// SIMATIC S7-200 project (STEP 7-Micro/WIN), CPU 224 CN REL 02.01

SYMBOL_TABLE USUARIO1
SF1              I0.0     // Sensor optico
SM3              I0.1     // Sensor magnetico de la Pinza
SM2              I0.2     // Sensor magnetico extendido cilindro horizontal
SM1              I0.3     // Sensor magnetico retraido cilindro horizontal
SM4              I0.4     // Sensor magnetico retraido cilindro de compresion
SM5              I0.5     // Sensor magnetico extendido cilindro de compresion
SB_2             I1.2     // Pulsador de paro
SB_1             I1.3     // Pulsador de marcha
QS               I1.4     // Zeta de emergencia
SA               I1.5     // Selector de modo
KV2              Q0.0     // Cilindro de la pinza
KV1              Q0.2     // Cilindro neumatico horizontal
KV3              Q0.3     // Cilindro neumatico de compresion
HL1              Q0.7     // Piloto indicador de parada
HL2              Q1.0     // Piloto indicador de marcha
HL3              Q1.1     // Piloto indicador de emergencia
E0               M0.0     // Estado 0
E1               M0.1     // Estado 1
E2               M0.2     // Estado 2
E3               M0.3     // Estado 3
E4               M0.4     // Estado 4
E5               M0.5     // Estado 5
E6               M0.6     // Estado 6
E7               M0.7     // Estado 7
EP               M1.0     // Estado de parada
EM               M1.1     // Estado de emergencia
END_SYMBOL_TABLE

ORGANIZATION_BLOCK PRINCIPAL:OB1
TITLE=COMENTARIOS DEL PROGRAMA
BEGIN
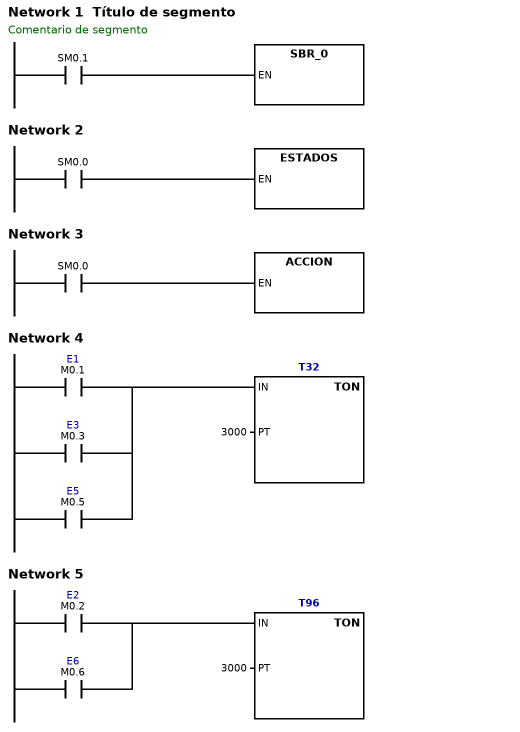
Network 1 // Título de segmento
// Comentario de segmento
LD     SM0.1
CALL   SBR_0:SBR0
Network 2
LD     SM0.0
CALL   ESTADOS:SBR1
Network 3
LD     SM0.0
CALL   ACCION:SBR2
Network 4
LD     E1:M0.1
O      E3:M0.3
O      E5:M0.5
TON    T32, 3000
Network 5
LD     E2:M0.2
O      E6:M0.6
TON    T96, 3000
END_ORGANIZATION_BLOCK

SUBROUTINE_BLOCK SBR_0:SBR0
TITLE=COMENTARIOS DE LA SUBRUTINA
BEGIN
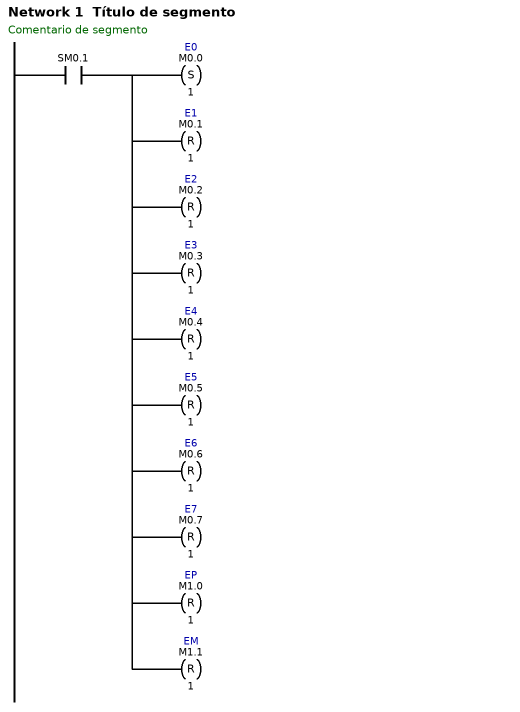
Network 1 // Título de segmento
// Comentario de segmento
LD     SM0.1
S      E0:M0.0, 1
R      E1:M0.1, 1
R      E2:M0.2, 1
R      E3:M0.3, 1
R      E4:M0.4, 1
R      E5:M0.5, 1
R      E6:M0.6, 1
R      E7:M0.7, 1
R      EP:M1.0, 1
R      EM:M1.1, 1
END_SUBROUTINE_BLOCK

SUBROUTINE_BLOCK ESTADOS:SBR1
TITLE=COMENTARIOS DE LA SUBRUTINA
BEGIN
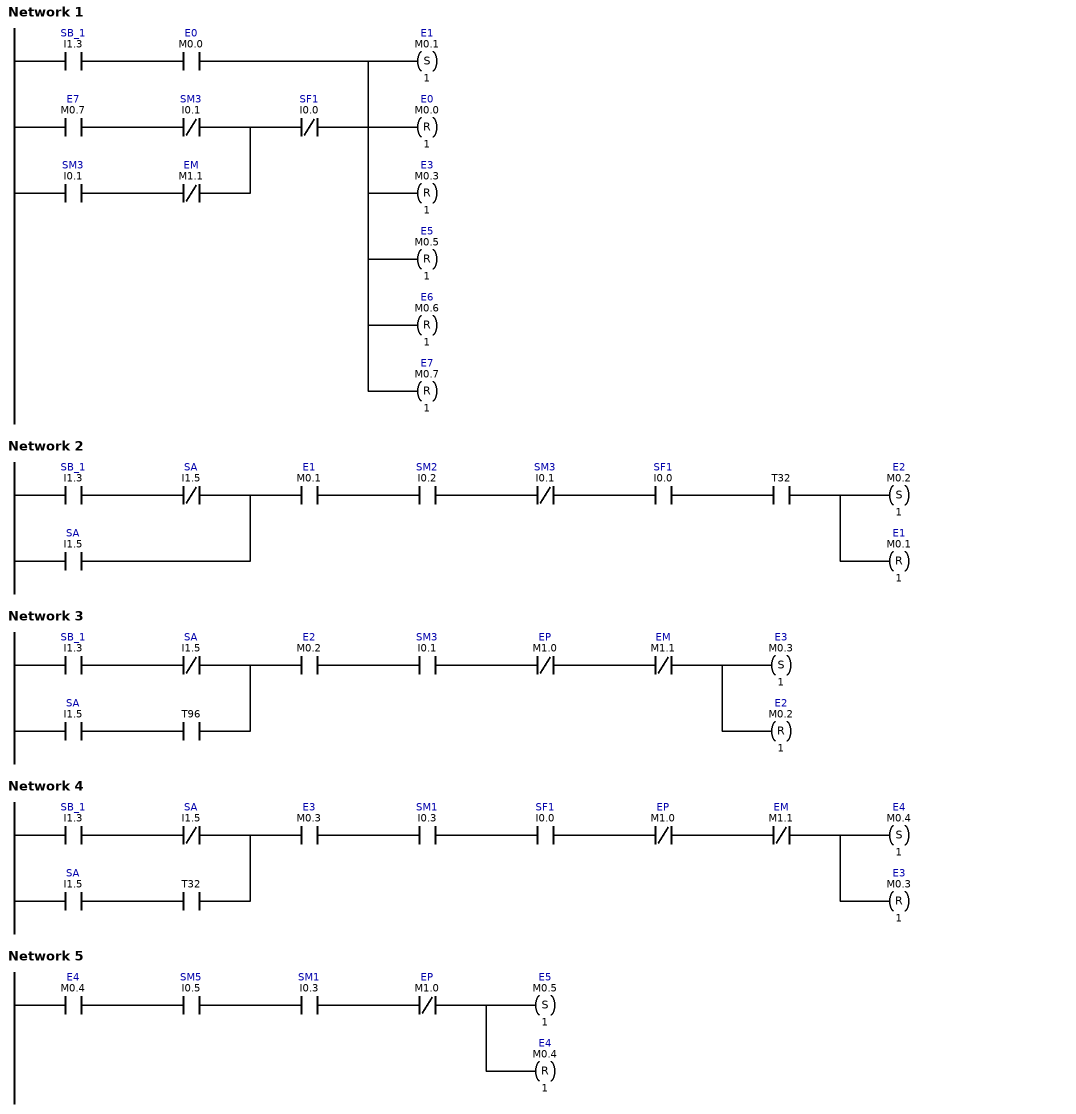
Network 1
LD     SB_1:I1.3
A      E0:M0.0
LD     E7:M0.7
AN     SM3:I0.1
LD     SM3:I0.1
AN     EM:M1.1
OLD
AN     SF1:I0.0
OLD
S      E1:M0.1, 1
R      E0:M0.0, 1
R      E3:M0.3, 1
R      E5:M0.5, 1
R      E6:M0.6, 1
R      E7:M0.7, 1
Network 2
LD     SB_1:I1.3
AN     SA:I1.5
O      SA:I1.5
A      E1:M0.1
A      SM2:I0.2
AN     SM3:I0.1
A      SF1:I0.0
A      T32
S      E2:M0.2, 1
R      E1:M0.1, 1
Network 3
LD     SB_1:I1.3
AN     SA:I1.5
LD     SA:I1.5
A      T96
OLD
A      E2:M0.2
A      SM3:I0.1
AN     EP:M1.0
AN     EM:M1.1
S      E3:M0.3, 1
R      E2:M0.2, 1
Network 4
LD     SB_1:I1.3
AN     SA:I1.5
LD     SA:I1.5
A      T32
OLD
A      E3:M0.3
A      SM1:I0.3
A      SF1:I0.0
AN     EP:M1.0
AN     EM:M1.1
S      E4:M0.4, 1
R      E3:M0.3, 1
Network 5
LD     E4:M0.4
A      SM5:I0.5
A      SM1:I0.3
AN     EP:M1.0
S      E5:M0.5, 1
R      E4:M0.4, 1
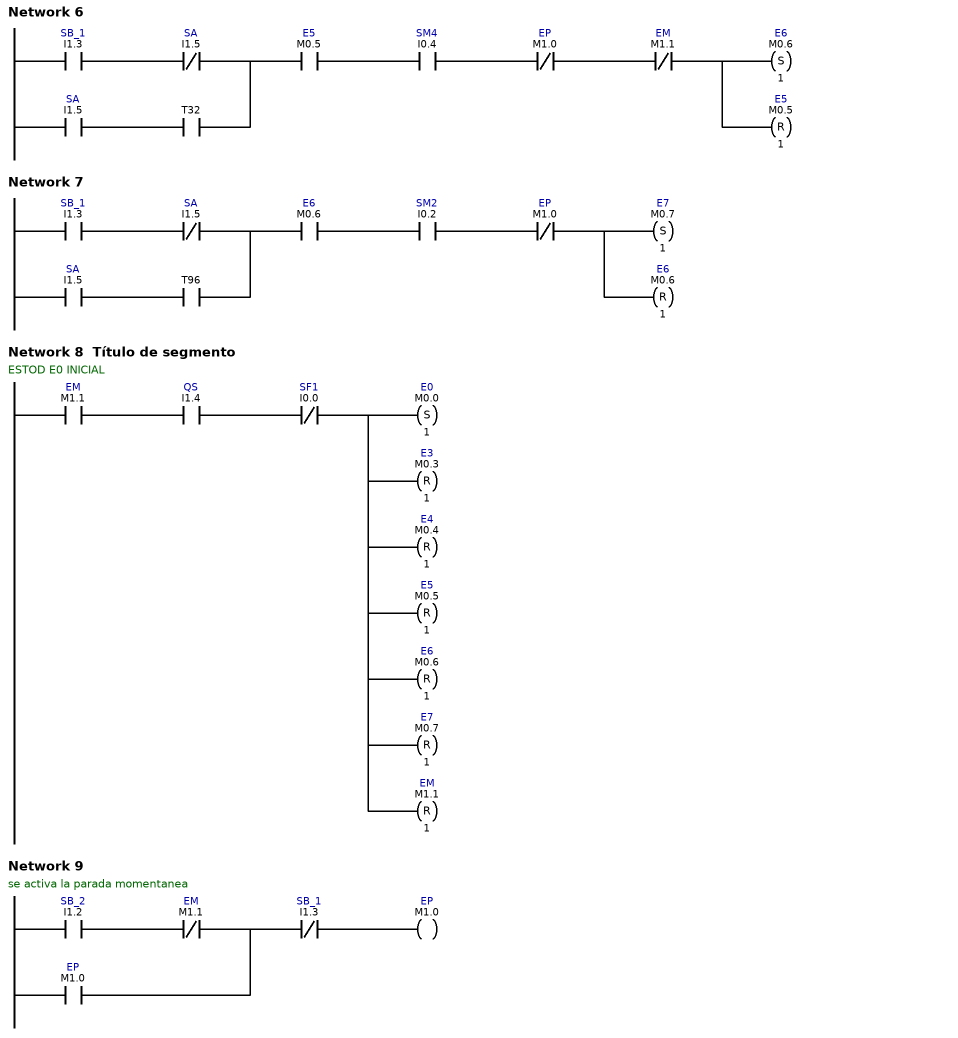
Network 6
LD     SB_1:I1.3
AN     SA:I1.5
LD     SA:I1.5
A      T32
OLD
A      E5:M0.5
A      SM4:I0.4
AN     EP:M1.0
AN     EM:M1.1
S      E6:M0.6, 1
R      E5:M0.5, 1
Network 7
LD     SB_1:I1.3
AN     SA:I1.5
LD     SA:I1.5
A      T96
OLD
A      E6:M0.6
A      SM2:I0.2
AN     EP:M1.0
S      E7:M0.7, 1
R      E6:M0.6, 1
Network 8 // Título de segmento
// ESTOD E0 INICIAL
LD     EM:M1.1
A      QS:I1.4
AN     SF1:I0.0
S      E0:M0.0, 1
R      E3:M0.3, 1
R      E4:M0.4, 1
R      E5:M0.5, 1
R      E6:M0.6, 1
R      E7:M0.7, 1
R      EM:M1.1, 1
Network 9
// se activa la parada momentanea
LD     SB_2:I1.2
AN     EM:M1.1
O      EP:M1.0
AN     SB_1:I1.3
=      EP:M1.0
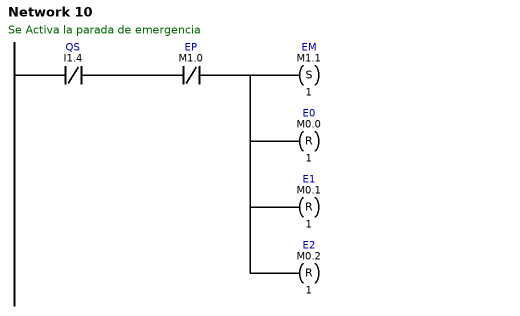
Network 10
// Se Activa la parada de emergencia
LDN    QS:I1.4
AN     EP:M1.0
S      EM:M1.1, 1
R      E0:M0.0, 1
R      E1:M0.1, 1
R      E2:M0.2, 1
END_SUBROUTINE_BLOCK

SUBROUTINE_BLOCK ACCION:SBR2
TITLE=COMENTARIOS DE LA SUBRUTINA
BEGIN
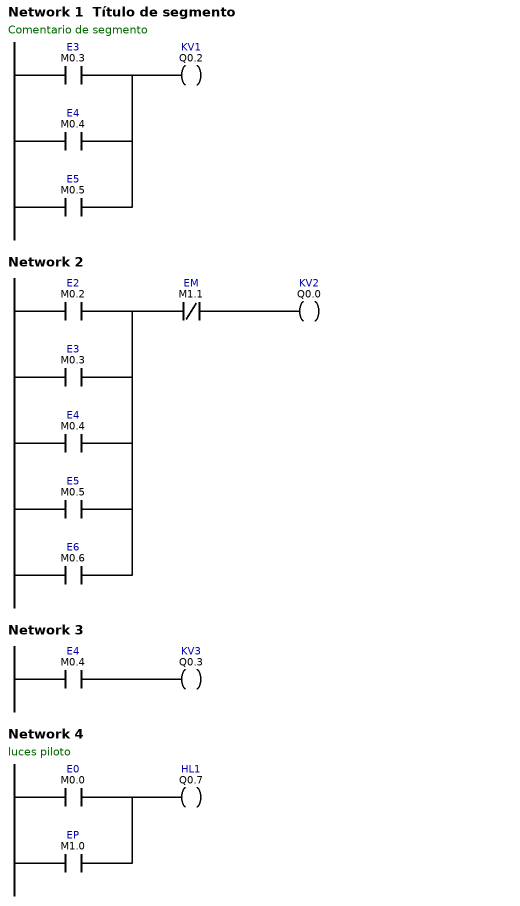
Network 1 // Título de segmento
// Comentario de segmento
LD     E3:M0.3
O      E4:M0.4
O      E5:M0.5
=      KV1:Q0.2
Network 2
LD     E2:M0.2
O      E3:M0.3
O      E4:M0.4
O      E5:M0.5
O      E6:M0.6
AN     EM:M1.1
=      KV2:Q0.0
Network 3
LD     E4:M0.4
=      KV3:Q0.3
Network 4
// luces piloto
LD     E0:M0.0
O      EP:M1.0
=      HL1:Q0.7
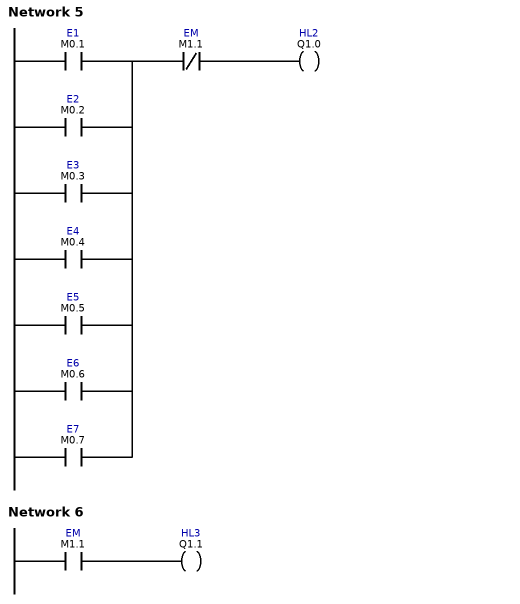
Network 5
LD     E1:M0.1
O      E2:M0.2
O      E3:M0.3
O      E4:M0.4
O      E5:M0.5
O      E6:M0.6
O      E7:M0.7
AN     EM:M1.1
=      HL2:Q1.0
Network 6
LD     EM:M1.1
=      HL3:Q1.1
END_SUBROUTINE_BLOCK
